Staubli VAL3: Algorithm6.pjx

--- Algorithm6.pjx ---
Parameters version=s8.10.5Cs9_BS2172 stackSize=5000 millimeterUnit=true
Program file=_CalpSphere.pgx
Program file=CalAdjustXY2.pgx
Program file=CalAdjustXY3.pgx
Program file=CalAdjustZ.pgx
Program file=CalToolPos3.pgx
Program file=CalToolPos4.pgx
Program file=CalToolPos7.pgx
Data file=Algorithm6.dtx
Library alias=matrix path=Disk://SmartTCP_CS9/MatrixLib/MatrixLib.pjx
Library alias=db path=Disk://SmartTCP_CS9/DataBase6/DataBase6.pjx

--- Algorithm6.dtx ---
public num nInverseMatrix1[4 4]
  [0,0] = 1.945193
  [0,1] = -1.712762
  [0,2] = 9.261268
  [1,0] = 0.502721
  [1,1] = 0.619141
  [1,2] = -1.663322
  [2,0] = 0.453432
  [2,1] = 1.0601144
  [2,2] = 3.220251
  [3,3] = 1
public num nMatrix1[4 4]
  [0,0] = 0.27407
  [0,1] = 1.118537
  [0,2] = -0.210464
  [1,0] = -0.17311
  [1,1] = 0.150611
  [1,2] = 0.575649
  [2,0] = 0.0183975
  [2,1] = -0.207079
  [2,2] = 0.150664
  [3,3] = 1
public num nMatrix2[4 4]
  [0,0] = 1
  [1,1] = 1
  [2,2] = 1
  [3,0] = 31.552388
  [3,1] = 103.369183
  [3,2] = -8.232965
  [3,3] = 1
public num nMatrix3[4 4]
  [0,0] = 1.945193
  [0,1] = -1.712762
  [0,2] = 9.261268
  [1,0] = 0.502721
  [1,1] = 0.619141
  [1,2] = -1.663322
  [2,0] = 0.453432
  [2,1] = 1.0601144
  [2,2] = 3.220251
  [3,0] = 109.608277
  [3,1] = 1.230419
  [3,2] = 93.766659
  [3,3] = 1
public num nTeach_3_1[4 4]
  [0,0] = -0.024705
  [0,1] = -0.0184623
  [0,2] = -0.999524
  [1,0] = -0.240476
  [1,1] = 0.970581
  [1,2] = -0.0119839
  [2,0] = 0.970341
  [2,1] = 0.240066
  [2,2] = -0.028418
  [3,0] = 888.833618
  [3,1] = -160.122184
  [3,2] = -41.507861
  [3,3] = 1
public num nTeach_3_2[4 4]
  [0,0] = -0.298775
  [0,1] = 0.518277
  [0,2] = -0.801326
  [1,0] = -0.0673661
  [1,1] = 0.82613
  [1,2] = 0.559438
  [2,0] = 0.951943
  [2,1] = 0.221128
  [2,2] = -0.211913
  [3,0] = 920.386007
  [3,1] = -217.720531
  [3,2] = -46.252531
  [3,3] = 1
public num nTeach_3_3[4 4]
  [0,0] = 0.130655
  [0,1] = -0.60026
  [0,2] = -0.789061
  [1,0] = -0.445377
  [1,1] = 0.67552
  [1,2] = -0.587633
  [2,0] = 0.885759
  [2,1] = 0.428207
  [2,2] = -0.179082
  [3,0] = 879.830904
  [3,1] = -114.351348
  [3,2] = -49.740826
  [3,3] = 1

--- _CalpSphere.pgx ---
program _CalpSphere(point x_p1, point x_p2, point x_p3, point x_p4, point& x_pCenter, bool& x_bStatus)
  local num x1
  local num x2
  local num x3
  local num x4
  local num y1
  local num y2
  local num y3
  local num y4
  local num z1
  local num z2
  local num z3
  local num z4
begin
  //球心算法
  x1=x_p1.trsf.x
  y1=x_p1.trsf.y
  z1=x_p1.trsf.z

  x2=x_p2.trsf.x
  y2=x_p2.trsf.y
  z2=x_p2.trsf.z

  x3=x_p3.trsf.x
  y3=x_p3.trsf.y
  z3=x_p3.trsf.z

  x4=x_p4.trsf.x
  y4=x_p4.trsf.y
  z4=x_p4.trsf.z

  //构造矩阵nMatrix1
  nMatrix1[0,0]=x2-x1
  nMatrix1[0,1]=x3-x1
  nMatrix1[0,2]=x4-x1
  nMatrix1[0,3]=0
  nMatrix1[1,0]=y2-y1
  nMatrix1[1,1]=y3-y1
  nMatrix1[1,2]=y4-y1
  nMatrix1[1,3]=0
  nMatrix1[2,0]=z2-z1
  nMatrix1[2,1]=z3-z1
  nMatrix1[2,2]=z4-z1
  nMatrix1[2,3]=0
  nMatrix1[3,0]=0
  nMatrix1[3,1]=0
  nMatrix1[3,2]=0
  nMatrix1[3,3]=1



  //构造矩阵nMatrix2
  nMatrix2[0,0]=1
  nMatrix2[0,1]=0
  nMatrix2[0,2]=0
  nMatrix2[0,3]=0

  nMatrix2[1,0]=0
  nMatrix2[1,1]=1
  nMatrix2[1,2]=0
  nMatrix2[1,3]=0

  nMatrix2[2,0]=0
  nMatrix2[2,1]=0
  nMatrix2[2,2]=1
  nMatrix2[2,3]=0

  nMatrix2[3,0]=(x2*x2+y2*y2+z2*z2-x1*x1-y1*y1-z1*z1)/2
  nMatrix2[3,1]=(x3*x3+y3*y3+z3*z3-x1*x1-y1*y1-z1*z1)/2
  nMatrix2[3,2]=(x4*x4+y4*y4+z4*z4-x1*x1-y1*y1-z1*z1)/2
  nMatrix2[3,3]=1

  call matrix:InverseMatrix(nMatrix1,nInverseMatrix1,x_bStatus)
  if x_bStatus==true
    //矩阵nMatrix1的逆矩阵nInverseMatrik1存在
    call matrix:MutliMatrix(nInverseMatrix1,nMatrix2,nMatrix3)
  endIf

  x_pCenter.trsf.x=nMatrix3[3,0]
  x_pCenter.trsf.y=nMatrix3[3,1]
  x_pCenter.trsf.z=nMatrix3[3,2]

end

--- CalAdjustXY2.pgx ---
public program CalAdjustXY2()
  local trsf l_trFlange
  local trsf l_trTCP
  local num x
  local num y
  local num z
begin
  //初始化数据
  l_trFlange={0,0,0,0,0,0}
  l_trTCP={0,0,0,0,0,0}
  //计算新的中心位置
  x=(db:pAdjustXY_2_1.trsf.x+db:pAdjustXY_2_2.trsf.x)/2
  y=(db:pAdjustXY_2_1.trsf.y+db:pAdjustXY_2_2.trsf.y)/2
  z=db:pAdjustXY_2_1.trsf.z
  //
  l_trFlange=db:pAdjustXY_2_1.trsf*!db:utCurrentTool.tValue.trsf
  if db:sMounting=="Floor"
    l_trTCP={x,y,z,0,180,0}
  elseIf db:sMounting=="Ceiling"
    l_trTCP={x,y,z,0,0,0}
  endIf
  db:tTool2.trsf=!l_trFlange*l_trTCP
  //
  db:tTool2.trsf.rx=db:tTool1.trsf.rx
  db:tTool2.trsf.ry=db:tTool1.trsf.ry
  db:tTool2.trsf.rz=db:tTool1.trsf.rz
  call db:hmiAlert("SaveInTool2","info")
end

--- CalAdjustXY3.pgx ---
public program CalAdjustXY3()
  local trsf l_trFlange
  local trsf l_trTCP
  local num x
  local num y
  local num z
begin
  l_trFlange={0,0,0,0,0,0}
  l_trTCP={0,0,0,0,0,0}
  x=db:pAdjustXY_3_2.trsf.x+db:pAdjustXY_3_3.trsf.x-db:pAdjustXY_3_1.trsf.x
  y=db:pAdjustXY_3_2.trsf.y+db:pAdjustXY_3_3.trsf.y-db:pAdjustXY_3_1.trsf.y
  z=db:pAdjustXY_3_1.trsf.z
  //
  l_trFlange=db:pAdjustXY_3_1.trsf*!db:utCurrentTool.tValue.trsf
  if db:sMounting=="Floor"
    l_trTCP={x,y,z,0,180,0}
  elseIf db:sMounting=="Ceiling"
    l_trTCP={x,y,z,0,0,0}
  endIf
  db:tTool2.trsf=!l_trFlange*l_trTCP
  //
  db:tTool2.trsf.rx=db:tTool1.trsf.rx
  db:tTool2.trsf.ry=db:tTool1.trsf.ry
  db:tTool2.trsf.rz=db:tTool1.trsf.rz
  call db:hmiAlert("SaveInTool2","info")
end

--- CalAdjustZ.pgx ---
public program CalAdjustZ()
  local num l_nDistance
  local trsf l_trZ
  local num l_nDir
begin
  l_nDistance=distance(db:pAdjustZ_2_1,db:pAdjustZ_2_2)
  switch db:sMounting
    case "Floor"
      l_nDir=1
    break
    case "Ceiling"
      l_nDir=-1
    break
    default
      l_nDir=1
    break
  endSwitch
  //
  if db:pAdjustZ_2_1.trsf.z<db:pAdjustZ_2_2.trsf.z
    l_trZ={0,0,-l_nDistance*l_nDir,0,0,0}
  else
    l_trZ={0,0,l_nDistance*l_nDir,0,0,0}
  endIf
  //
  db:tTool3.trsf=db:utCurrentTool.tValue.trsf*l_trZ
  db:tTool3.trsf.rx=db:tTool1.trsf.rx
  db:tTool3.trsf.ry=db:tTool1.trsf.ry
  db:tTool3.trsf.rz=db:tTool1.trsf.rz
  call db:hmiAlert("SaveInTool3","info")
end

--- CalToolPos3.pgx ---
public program CalToolPos3(tool& x_tTool)
  local num ax1
  local num ax2
  local num ax3
  local num ay1
  local num ay2
  local num ay3
  local num az1
  local num az2
  local num az3
  local bool l_bStatus
  local pointRx l_p1
  local pointRx l_p2
  local pointRx l_p3
  local point l_pCenter
  local trsf l_trP1
  local trsf l_trP2
  local trsf l_trP3
  local num nx1
  local num nx2
  local num nx3
  local num ny1
  local num ny2
  local num ny3
  local num nz1
  local num nz2
  local num nz3
  local num ox1
  local num ox2
  local num ox3
  local num oy1
  local num oy2
  local num oy3
  local num oz1
  local num oz2
  local num oz3
  local num xf1
  local num xf2
  local num xf3
  local num yf1
  local num yf2
  local num yf3
  local num zf1
  local num zf2
  local num zf3
begin
  //3个带姿态的点求工具值XYZ
  l_trP1=db:pTeach1.trsf
  l_trP2=db:pTeach2.trsf
  l_trP3=db:pTeach3.trsf
  //
  //pTeach_3_1转成矩阵nTeach_3_1
  call matrix:Trsf2Matrix(l_trP1,nTeach_3_1)
  //pTeach_3_2转成矩阵nTeach_3_2
  call matrix:Trsf2Matrix(l_trP2,nTeach_3_2)
  //pTeach_3_3转成矩阵nTeach_3_3
  call matrix:Trsf2Matrix(l_trP3,nTeach_3_3)
  //
  //分解矩阵nTeach_3_1
  nx1=nTeach_3_1[0,0]
  ny1=nTeach_3_1[0,1]
  nz1=nTeach_3_1[0,2]
  ox1=nTeach_3_1[1,0]
  oy1=nTeach_3_1[1,1]
  oz1=nTeach_3_1[1,2]
  ax1=nTeach_3_1[2,0]
  ay1=nTeach_3_1[2,1]
  az1=nTeach_3_1[2,2]
  xf1=nTeach_3_1[3,0]
  yf1=nTeach_3_1[3,1]
  zf1=nTeach_3_1[3,2]
  //
  //分解矩阵nTeach_3_2
  nx2=nTeach_3_2[0,0]
  ny2=nTeach_3_2[0,1]
  nz2=nTeach_3_2[0,2]
  ox2=nTeach_3_2[1,0]
  oy2=nTeach_3_2[1,1]
  oz2=nTeach_3_2[1,2]
  ax2=nTeach_3_2[2,0]
  ay2=nTeach_3_2[2,1]
  az2=nTeach_3_2[2,2]
  xf2=nTeach_3_2[3,0]
  yf2=nTeach_3_2[3,1]
  zf2=nTeach_3_2[3,2]
  //
  //分解矩阵nTeach_3_3
  nx3=nTeach_3_3[0,0]
  ny3=nTeach_3_3[0,1]
  nz3=nTeach_3_3[0,2]
  ox3=nTeach_3_3[1,0]
  oy3=nTeach_3_3[1,1]
  oz3=nTeach_3_3[1,2]
  ax3=nTeach_3_3[2,0]
  ay3=nTeach_3_3[2,1]
  az3=nTeach_3_3[2,2]
  xf3=nTeach_3_3[3,0]
  yf3=nTeach_3_3[3,1]
  zf3=nTeach_3_3[3,2]
  //
  //***************************************************************************************
  //  │nx1-nx2 , ox1-ox2 , ax1-ax2 ,   0  │   │1 , 0 , 0, Tx│   │1 , 0 , 0, xf2-xf1│
  //  │ny2-ny3 , oy2-oy3 , ay2-ay3 ,   0  │ * │0 , 1 , 0, Ty│ = │0 , 1 , 0, yf3-yf2│
  //  │nz1-nz3 , oz1-oz3 , az1-az3 ,   0  │   │0 , 0 , 1, Tz│   │0 , 0 , 1, zf3-zf1│
  //  │   0    ,    0    ,    0    ,   1  │   │0 , 0 , 0,  1│   │0 , 0 , 0,    1   │
  //***************************************************************************************
  //构造矩阵nMatrix1
  nMatrix1[0,0]=nx1-nx2
  nMatrix1[0,1]=ny2-ny3
  nMatrix1[0,2]=nz1-nz3
  nMatrix1[0,3]=0
  nMatrix1[1,0]=ox1-ox2
  nMatrix1[1,1]=oy2-oy3
  nMatrix1[1,2]=oz1-oz3
  nMatrix1[1,3]=0
  nMatrix1[2,0]=ax1-ax2
  nMatrix1[2,1]=ay2-ay3
  nMatrix1[2,2]=az1-az3
  nMatrix1[2,3]=0
  nMatrix1[3,0]=0
  nMatrix1[3,1]=0
  nMatrix1[3,2]=0
  nMatrix1[3,3]=1

  //构造矩阵nMatrix2
  nMatrix2[0,0]=1
  nMatrix2[0,1]=0
  nMatrix2[0,2]=0
  nMatrix2[0,3]=0

  nMatrix2[1,0]=0
  nMatrix2[1,1]=1
  nMatrix2[1,2]=0
  nMatrix2[1,3]=0

  nMatrix2[2,0]=0
  nMatrix2[2,1]=0
  nMatrix2[2,2]=1
  nMatrix2[2,3]=0

  nMatrix2[3,0]=xf2-xf1
  nMatrix2[3,1]=yf3-yf2
  nMatrix2[3,2]=zf3-zf1
  nMatrix2[3,3]=1
  //***************************************************************************************
  call matrix:InverseMatrix(nMatrix1,nInverseMatrix1,l_bStatus)
  if l_bStatus==false
    //如果nMatrix1不可逆则需重新示教点
    call db:hmiAlert("DeviationIsTooLarge","warning")
  else
    call matrix:MutliMatrix(nInverseMatrix1,nMatrix2,nMatrix3)

    x_tTool.trsf.x=nMatrix3[3,0]
    x_tTool.trsf.y=nMatrix3[3,1]
    x_tTool.trsf.z=nMatrix3[3,2]
    x_tTool.trsf.rx=0
    x_tTool.trsf.ry=0
    x_tTool.trsf.rz=0
  endIf
  //定义中心点xyz
  l_pCenter.trsf=l_p1.trsf*x_tTool.trsf
  //定义中心点RxRyRz
  if db:sMounting=="Floor"
    l_pCenter.trsf.rx=0
    l_pCenter.trsf.ry=180
    l_pCenter.trsf.rz=0
  elseIf db:sMounting=="Ceiling"
    l_pCenter.trsf.rx=0
    l_pCenter.trsf.ry=0
    l_pCenter.trsf.rz=0
  endIf
  x_tTool.trsf=!l_p1.trsf*l_pCenter.trsf
  call db:hmiAlert("SaveInTool1","info")
end

--- CalToolPos4.pgx ---
public program CalToolPos4(tool& x_tTool)
  local bool l_bStatus
  local pointRx l_p1
  local pointRx l_p2
  local pointRx l_p3
  local pointRx l_p4
  local point l_pCenter
  local tool l_t1
  local tool l_t2
  local tool l_t3
  local tool l_t4
  local num x1
  local num x2
  local num x3
  local num x4
  local num y1
  local num y2
  local num y3
  local num y4
  local num z1
  local num z2
  local num z3
  local num z4
begin
  //取中心点xyz
  l_p1=db:pTeach1
  l_p2=db:pTeach2
  l_p3=db:pTeach3
  l_p4=db:pTeach4
  l_pCenter=here(flange,world)
  call _CalpSphere(l_p1,l_p2,l_p3,l_p4,l_pCenter,l_bStatus)

  if l_bStatus==false
    call db:hmiAlert("DeviationIsTooLarge","warning")
  else
    if db:sMounting=="Floor"
      l_pCenter.trsf.rx=0
      l_pCenter.trsf.ry=180
      l_pCenter.trsf.rz=0
    elseIf db:sMounting=="Ceiling"
      l_pCenter.trsf.rx=0
      l_pCenter.trsf.ry=0
      l_pCenter.trsf.rz=0
    endIf
    l_t1.trsf=!l_p1.trsf*l_pCenter.trsf
    l_t2.trsf=!l_p2.trsf*l_pCenter.trsf
    l_t3.trsf=!l_p3.trsf*l_pCenter.trsf
    l_t4.trsf=!l_p4.trsf*l_pCenter.trsf
    x_tTool.trsf.x=(l_t1.trsf.x+l_t2.trsf.x+l_t3.trsf.x+l_t4.trsf.x)/4
    x_tTool.trsf.y=(l_t1.trsf.y+l_t2.trsf.y+l_t3.trsf.y+l_t4.trsf.y)/4
    x_tTool.trsf.z=(l_t1.trsf.z+l_t2.trsf.z+l_t3.trsf.z+l_t4.trsf.z)/4
    x_tTool.trsf.rx=l_t1.trsf.rx
    x_tTool.trsf.ry=l_t1.trsf.ry
    x_tTool.trsf.rz=l_t1.trsf.rz
    call db:hmiAlert("SaveInTool1","info")
  endIf
end

--- CalToolPos7.pgx ---
public program CalToolPos7(tool& x_tTool)
  local frame l_fFrame
  local num l_nFrameErr
  local point l_pCenter
  local bool l_bStatus
  local point l_p5flange
begin
  //定义中心点xyz
  link(l_fFrame,world)
  link(l_pCenter,world)
  //
  call _CalpSphere(db:pTeach1,db:pTeach2,db:pTeach3,db:pTeach4,l_pCenter,l_bStatus)
  l_nFrameErr=setFrame(db:pTeach5,db:pTeach6,db:pTeach7,l_fFrame)
  switch l_nFrameErr
    case 0
      l_pCenter.trsf.rx=l_fFrame.trsf.rx
      l_pCenter.trsf.ry=l_fFrame.trsf.ry
      l_pCenter.trsf.rz=l_fFrame.trsf.rz
      x_tTool.trsf=!db:pTeach5.trsf*l_pCenter.trsf
    break
    case -1,-2
      call db:hmiAlert("DeviationIsTooLarge","warning")
    break
  endSwitch
  call db:hmiAlert("SaveInTool1","info")
end
